# B&R Automation Studio project ProjetoFinalRobotica
Automation Studio 4.1.14.40 SP

## Configuration Config1

CPU 4PP481.1043-B5, AutomationRuntime E3.10, Build 4.1.2, Vc V4.15.9

### Task classes (Cpu.sw)
```
Cyclic#1 (cycle 10000 us, tolerance 10000 us):
  NewProgram <- NewProgram.prg
VcDataObjects: Visu <- Visualisation.Visu.dob
Binaries: arial, Visu02, vccovl, vcdsloc, vcfntttf, vcbclass, vcrt, Visu03, vcfile, vcdsint, vccbtn, vcgclass, vcpdsw, vcshared, vcalarm, arialbd, vcpfpp30, vcmgr, vcpdpp30, Visu01, vctcal, vcpk, vcpfmtcx, vcptelo, ashwd, sysconf, asfw, arconfig, iomap, arialxsr, vcctrend, vccline, vccshape, vccbmp, vcclbox, vccalarm, vccstr, vcchspot, vccgauge, vccurl, vccslider, vccnum, vccdt, vcxml, vccbar, vcchtml, vcctext
Libraries: standard, dataobj, vcresman, fileio, astime, asieccon, AsUDP, Runtime
```

### Hardware
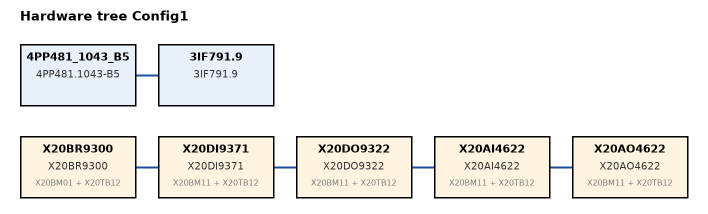
```
3IF791.9 : 3IF791.9 v1.0.0.1  [SS -> 4PP481_1043_B5.SS1]
4PP481_1043_B5 : 4PP481.1043-B5 v1.0.0.0
  Connector IF5:
    ActivateDevice = 1
    Mode = Manual
    InternetAddress = 192.168.0.70
  Cyclic1Duration = 10000
  Cyclic1Tolerance = 10000
  Cyclic2Duration = 20000
  Cyclic2Tolerance = 20000
  Cyclic3Duration = 50000
  Cyclic3Tolerance = 50000
  Cyclic4Duration = 100000
  Cyclic4Tolerance = 100000
  Cyclic5Duration = 200000
  Cyclic5Tolerance = 200000
  Cyclic6Duration = 500000
  Cyclic6Tolerance = 500000
  Cyclic7Duration = 1000000
  Cyclic7Tolerance = 1000000
  Cyclic8Duration = 10000
  Cyclic8Tolerance = 30000000
  VcObjectName = Visu
  KeyMappingFile = VC\4PP481_1043_B5.dis
X20AI4622 : X20AI4622 v1.0.2.0  [SS1 -> X20TB12c.SS; SL -> X20BM11b.SL1]
X20AO4622 : X20AO4622 v1.0.4.0  [SS1 -> X20TB12e.SS; SL -> X20BM11c.SL1]
X20BM01 : X20BM01 v1.0.0.1
X20BM11 : X20BM11 v1.0.0.0  [X2X1 -> X20BM01.X2X2]
X20BM11a : X20BM11 v1.0.0.0  [X2X1 -> X20BM11.X2X2]
X20BM11b : X20BM11 v1.0.0.0  [X2X1 -> X20BM11a.X2X2]
X20BM11c : X20BM11 v1.0.0.0  [X2X1 -> X20BM11b.X2X2]
X20BR9300 : X20BR9300 v1.0.2.4  [SS1 -> X20TB12.SS; SL -> X20BM01.SL1; X2X1 -> 3IF791.9.IF1]
X20DI9371 : X20DI9371 v1.0.1.1  [SS1 -> X20TB12a.SS; SL -> X20BM11.SL1]
X20DO9322 : X20DO9322 v1.0.2.2  [SS1 -> X20TB12b.SS; SL -> X20BM11a.SL1]
X20TB12 : X20TB12 v1.0.0.0
X20TB12a : X20TB12 v1.0.0.0
X20TB12b : X20TB12 v1.0.0.0
X20TB12c : X20TB12 v1.0.0.0
X20TB12e : X20TB12 v1.0.0.0
```

### IoMap.iom - 4PP481_1043_B5/IoMap.iom
```iecst
(********************************************************************
 * COPYRIGHT --
 ********************************************************************
 * File: IoMap.iom
 * Author: supervisorio
 * Created: February 20, 2025
 ********************************************************************
 * IO mapping file
 ********************************************************************)
VAR_CONFIG
	::NewProgram:Jaka_DI3 AT %QX."X20DO9322".DigitalOutput01;
	::NewProgram:Jaka_DI2 AT %QX."X20DO9322".DigitalOutput02;
	::NewProgram:Jaka_DI1 AT %QX."X20DO9322".DigitalOutput03;
	::NewProgram:Staubli_DI12 AT %QX."X20DO9322".DigitalOutput05;
	::NewProgram:Staubli_DI13 AT %QX."X20DO9322".DigitalOutput06;
	::NewProgram:Staubli_DI14 AT %QX."X20DO9322".DigitalOutput07;
	::NewProgram:Staubli_DI15 AT %QX."X20DO9322".DigitalOutput08;
	::NewProgram:Esteira_StaubliJaka AT %QX."X20DO9322".DigitalOutput11;
	::NewProgram:Esteira_JakaStaubli AT %QX."X20DO9322".DigitalOutput12;
	::NewProgram:Jaka_DO7 AT %IX."X20DI9371".DigitalInput01;
	::NewProgram:Jaka_DO6 AT %IX."X20DI9371".DigitalInput02;
	::NewProgram:Jaka_DO5 AT %IX."X20DI9371".DigitalInput03;
	::NewProgram:Staubli_DO4 AT %IX."X20DI9371".DigitalInput05;
	::NewProgram:Staubli_DO5 AT %IX."X20DI9371".DigitalInput06;
	::NewProgram:Staubli_DO6 AT %IX."X20DI9371".DigitalInput07;
	::NewProgram:Staubli_DO7 AT %IX."X20DI9371".DigitalInput08;
	::NewProgram:Sensor_Staubli AT %IX."X20DI9371".DigitalInput09;
	::NewProgram:Sensor_Jaka AT %IX."X20DI9371".DigitalInput10;
	::NewProgram:Emergencia AT %IX."X20DI9371".DigitalInput12;
END_VAR
```

## Logical view

Binary libraries used (declarations not repeated): operator, runtime, astime, AsIecCon, standard, AsUDP

### Global.typ - Global data types
```iecst
(********************************************************************
 * COPYRIGHT --
 ********************************************************************
 * File: Global.typ
 * Author: supervisorio
 * Created: February 20, 2025
 ********************************************************************
 * Global data types of project CLP_ROBO
 ********************************************************************)

TYPE
	feeder_status_typ : 	STRUCT
		power : BOOL;
		home : BOOL;
		axisErrorNumber : UINT;
		axisErrorText : STRING[255];
	END_STRUCT;
	feeder_cmd_typ : 	STRUCT
		requestToPut : BOOL;
	END_STRUCT;
	feeder_typ : 	STRUCT
		cmd : feeder_cmd_typ;
		status : feeder_status_typ;
	END_STRUCT;
	main_status_money_typ : 	STRUCT
		changedMoney : REAL;
		cent1 : USINT;
		cent2 : USINT;
		cent5 : USINT;
		cent10 : USINT;
		cent20 : USINT;
		cent50 : USINT;
		euro1 : UDINT;
		euro2 : UDINT;
	END_STRUCT;
	main_status_progress_typ : 	STRUCT
		total : REAL;
		current : REAL;
	END_STRUCT;
	main_status_typ : 	STRUCT
		money : main_status_money_typ;
		progressStep : USINT;
		curPage : UINT;
		curLanguage : UINT;
		startProgressStep : USINT;
	END_STRUCT;
	main_par_recipe_typ : 	STRUCT
		price : REAL;
		setTemp : REAL;
		milk : REAL;
		sugar : REAL;
		coffee : REAL;
		water : REAL;
	END_STRUCT;
	main_par_typ : 	STRUCT
		coffeeType : SINT;
		givenMoney : REAL;
		recipe : main_par_recipe_typ;
	END_STRUCT;
	main_cmd_typ : 	STRUCT
		switchOnOff : BOOL;
		errorAck : BOOL;
		start : BOOL;
		vis : main_cmd_vis_typ;
	END_STRUCT;
	main_cmd_vis_typ : 	STRUCT
		newPage : UINT;
		startFlag : BOOL;
		startButtonColor : UINT;
		waterTempColor : UINT;
		messageColor : UINT;
		messageIndex : USINT;
		euro2hidden : UINT;
		euro1hidden : UINT;
		cent50hidden : UINT;
		cent20hidden : UINT;
		cent10hidden : UINT;
		cent5hidden : UINT;
		cent2hidden : UINT;
		cent1hidden : UINT;
		newLanguage : UINT;
	END_STRUCT;
	main_typ : 	STRUCT
		cmd : main_cmd_typ;
		par : main_par_typ;
		status : main_status_typ;
	END_STRUCT;
	conveyor_typ : 	STRUCT
		status : conveyor_status_typ;
	END_STRUCT;
	conveyor_status_typ : 	STRUCT
		power : BOOL;
		home : BOOL;
		axisErrorNumber : UINT;
		axisErrorText : STRING[255];
		readyToTake : BOOL;
	END_STRUCT;
	brewing_par_typ : 	STRUCT
		coffeeType : USINT;
	END_STRUCT;
	brewing_cmd_typ : 	STRUCT
		start : BOOL;
	END_STRUCT;
	brewing_status_typ : 	STRUCT
		done : BOOL;
		sBrewingStep : UINT;
		brewingStepText : STRING[64];
	END_STRUCT;
	brewing_typ : 	STRUCT
		cmd : brewing_cmd_typ;
		par : brewing_par_typ;
		status : brewing_status_typ;
	END_STRUCT;
	heating_status_typ : 	STRUCT
		setTempOK : BOOL;
		actTemp : REAL;
	END_STRUCT;
	heating_cmd_typ : 	STRUCT
		start : BOOL;
		updatePIDpar : BOOL;
	END_STRUCT;
	heating_typ : 	STRUCT
		cmd : heating_cmd_typ;
		status : heating_status_typ;
	END_STRUCT;
END_TYPE
```

### Package Logical/Libraries - Global libraries

- Visualisation Logical/Visualisation (not shown)

### Program Logical/NewProgram (IEC) - Program

#### NewProgramCyclic.st - Cyclic code
```iecst
(********************************************************************
 * COPYRIGHT --
 ********************************************************************
 * PROGRAM: NewProgram
 * File: NewProgramCyclic.st
 * Author: supervisorio
 * Created: May 29, 2026
 ********************************************************************
 * Whiteboard application (docs/whiteboard-application.md):
 *   1. Jaka puts the plate (NUM_PECAS parts in its holes) on the conveyor.
 *   2. The conveyor brings the plate TO the Staubli.
 *   3. Staubli puts the plate on its table AND the parts on the board.
 *   4. Staubli picks the marker from its table, draws a square around
 *      each part AND puts the marker back.
 * NUM_PECAS (NewProgram.var) is 1 FOR now: one part, one square.
 * Every robot task uses a four-phase handshake (no timers):
 *   PLC sets CMD -> robot sets DONE -> PLC clears CMD -> robot clears DONE.
 * One run per press OF the start button: Ligar is cleared at the end
 * OF the cycle AND on E-stop.
 ********************************************************************)
PROGRAM _CYCLIC

	TmrPulso(IN := Ligar AND Emergencia, PT := T#1s);
	TmrDI12(IN := Etapa = 2, PT := T#1s);

	IF Ligar AND Emergencia THEN

		Jaka_DI2 := NOT TmrPulso.Q;		//Pulse: ON for the first 1 s of the cycle, then OFF
		Staubli_DI13 := NOT TmrPulso.Q;
		LIGA_JAKA := TRUE;

		CASE Etapa OF

			0: (* Start *)
				PlacaNaEsteira := FALSE;
				PlacaChegou := FALSE;
				PecasNoQuadro := FALSE;
				CicloConcluido := FALSE;
				iPecasNoQuadro := 0;
				iQuadrados := 0;
				iTempoCiclo_s := 0;
				Jaka_DI3 := TRUE;						//CMD Jaka: put the plate on the conveyor
				Etapa := 1;

			1: (* Plate to the Staubli *)
				IF Jaka_DO7 = TRUE THEN
					//Jaka_DI3 := FALSE;					//Jaka done: plate on the conveyor
					PlacaNaEsteira := TRUE;
					Esteira_JakaStaubli := TRUE;
					Jaka_DI2 := FALSE;	//Carry the plate to the Staubli
				END_IF;

				IF Esteira_JakaStaubli AND Sensor_Staubli THEN
					Esteira_JakaStaubli := FALSE;		//Plate arrived
					PlacaChegou := TRUE;
				END_IF;

				//Wait for the Jaka to clear DONE
				IF PlacaChegou AND NOT Jaka_DO7 THEN
					Etapa := 2;
				END_IF;

			2: (* Staubli: plate on the table, parts on the board *)
				Staubli_DI12 := NOT TmrDI12.Q;			//CMD Staubli: plate to the table, parts to the board
				IF Staubli_DO4 THEN
					Staubli_DI12 := FALSE;				//Staubli done: parts on the board
					PecasNoQuadro := TRUE;
					iPecasNoQuadro := NUM_PECAS;
					Etapa := 3;
				END_IF;

			3: (* Wait for the Staubli to clear DONE *)
				IF NOT Staubli_DO4 THEN
					Etapa := 4;
				END_IF;

			4: (* Staubli: pick the marker, draw the squares, put the marker back *)
				Staubli_DI14 := TRUE;					//CMD Staubli: pick the marker and draw
				IF Staubli_DO5 THEN
					Staubli_DI14 := FALSE;				//Staubli done: squares drawn, marker stored
					iQuadrados := NUM_PECAS;
					Etapa := 5;
				END_IF;

			5: (* Finish: wait for the Staubli to clear DONE *)
				IF NOT Staubli_DO5 THEN
					iContador := iContador + 1;			//Completed cycles
					CicloConcluido := TRUE;
					Ligar := FALSE;						//One run per start; press Ligar again for the next
					Etapa := 0;
				END_IF;

		END_CASE;

	ELSE
		//Stop or E-stop: every command and enable goes FALS
		LIGA_JAKA := FALSE;
		Jaka_DI1 := FALSE;
		Jaka_DI2 := FALSE;
		Jaka_DI3 := FALSE;
		Staubli_DI12 := FALSE;
		Staubli_DI13 := FALSE;
		Staubli_DI14 := FALSE;
		Staubli_DI15 := FALSE;
		Esteira_JakaStaubli := FALSE;
		Esteira_StaubliJaka := FALSE;
		IF NOT Emergencia THEN
			Ligar := FALSE;							//Releasing the E-stop must not restart the cell
		END_IF;
		Etapa := 0;

		//Reset the process state too, so the HMI colors, counters and progress go back to "waiting".
		//Skipped right after a finished cycle: CicloConcluido stays TRUE until the next start,
		//so the "done" state and the cycle time stay on screen.
		IF NOT CicloConcluido THEN
			PlacaNaEsteira := FALSE;
			PlacaChegou := FALSE;
			PecasNoQuadro := FALSE;
			iPecasNoQuadro := 0;
			iQuadrados := 0;
			iTempoCiclo_s := 0;
		END_IF;
	END_IF;

	//Progress counters from the robots' optional pulses (Staubli DO6 = part placed, DO7 = square drawn)
	PulsoPeca(CLK := Staubli_DO6);
	IF PulsoPeca.Q AND Etapa = 2 AND iPecasNoQuadro < NUM_PECAS THEN
		iPecasNoQuadro := iPecasNoQuadro + 1;
	END_IF;
	PulsoQuadrado(CLK := Staubli_DO7);
	IF PulsoQuadrado.Q AND Etapa = 4 AND iQuadrados < NUM_PECAS THEN
		iQuadrados := iQuadrados + 1;
	END_IF;

	//Cycle time (kept on screen after the cycle ends)
	TempoCiclo(IN := Etapa > 0, PT := T#30m);
	IF Etapa > 0 THEN
		iTempoCiclo_s := DINT_TO_INT(TIME_TO_DINT(TempoCiclo.ET) / 1000);
	END_IF;

	//Where the plate is: 0 = Jaka, 1 = conveyor, 2 = Staubli
	IF PlacaChegou THEN
		iPlaca := 2;
	ELSIF PlacaNaEsteira THEN
		iPlaca := 1;
	ELSE
		iPlaca := 0;
	END_IF;

	//HMI colors (palette index): COR_ESPERA = waiting, COR_ANDAMENTO = running, COR_FEITO = done
	IF PlacaNaEsteira THEN iCorJaka := COR_FEITO; ELSIF Jaka_DI3 THEN iCorJaka := COR_ANDAMENTO; ELSE iCorJaka := COR_ESPERA; END_IF;
	IF PlacaChegou THEN iCorEsteira := COR_FEITO; ELSIF Esteira_JakaStaubli THEN iCorEsteira := COR_ANDAMENTO; ELSE iCorEsteira := COR_ESPERA; END_IF;
	IF PecasNoQuadro THEN iCorPecas := COR_FEITO; ELSIF Staubli_DI12 THEN iCorPecas := COR_ANDAMENTO; ELSE iCorPecas := COR_ESPERA; END_IF;
	IF CicloConcluido OR Etapa = 5 THEN iCorDesenho := COR_FEITO; ELSIF Etapa = 4 THEN iCorDesenho := COR_ANDAMENTO; ELSE iCorDesenho := COR_ESPERA; END_IF;
	IF CicloConcluido THEN iCorConcluido := COR_FEITO; ELSIF Etapa = 5 THEN iCorConcluido := COR_ANDAMENTO; ELSE iCorConcluido := COR_ESPERA; END_IF;

	//Whiteboard (one part and its square on the HMI)
	IF iPecasNoQuadro >= 1 THEN iCorPeca := COR_PECA; ELSE iCorPeca := COR_VAZIO; END_IF;
	IF iQuadrados >= 1 THEN iCorQuadrado := COR_TINTA; ELSE iCorQuadrado := COR_QUADRO; END_IF;

	IF iPlaca = 0 THEN iCorPlacaJaka := COR_FEITO; ELSE iCorPlacaJaka := COR_ESPERA; END_IF;
	IF iPlaca = 1 THEN iCorPlacaEsteira := COR_FEITO; ELSE iCorPlacaEsteira := COR_ESPERA; END_IF;
	IF iPlaca = 2 THEN iCorPlacaStaubli := COR_FEITO; ELSE iCorPlacaStaubli := COR_ESPERA; END_IF;

	iProgresso := iPecasNoQuadro + iQuadrados;	//0..2*NUM_PECAS on the progress bar

	//Digital twin: send the I/O state to the bridge PC (TwinSender.st)
	TwinSender;

END_PROGRAM
```

#### TwinSender.st - Digital twin UDP sender (action)
```iecst
(********************************************************************
 * COPYRIGHT --
 ********************************************************************
 * Program: NewProgram
 * File: TwinSender.st
 ********************************************************************
 * Digital twin: sends the I/O state to the bridge PC over UDP.
 * Called once per scan at the end of _CYCLIC.
 * Packet layout: docs/publishing-plan/02-plc-udp-sender.md
 * Needs the AsUDP library (Logical View > Libraries > Add Object).
 * Send errors are only counted: the cell must never depend on the
 * bridge PC being present.
 ********************************************************************)
ACTION TwinSender:

	(* Bytes 0..11: X20DI9371 channels 1..12 *)
	TwinPacket[0]  := BOOL_TO_USINT(Jaka_DO7);
	TwinPacket[1]  := BOOL_TO_USINT(Jaka_DO6);
	TwinPacket[2]  := BOOL_TO_USINT(Jaka_DO5);
	TwinPacket[4]  := BOOL_TO_USINT(Staubli_DO4);
	TwinPacket[5]  := BOOL_TO_USINT(Staubli_DO5);
	TwinPacket[6]  := BOOL_TO_USINT(Staubli_DO6);
	TwinPacket[7]  := BOOL_TO_USINT(Staubli_DO7);
	TwinPacket[8]  := BOOL_TO_USINT(Sensor_Staubli);
	TwinPacket[9]  := BOOL_TO_USINT(Sensor_Jaka);
	TwinPacket[11] := BOOL_TO_USINT(Emergencia);

	(* Bytes 12..23: X20DO9322 channels 1..12 *)
	TwinPacket[12] := BOOL_TO_USINT(Jaka_DI3);
	TwinPacket[13] := BOOL_TO_USINT(LIGA_JAKA);
	TwinPacket[14] := BOOL_TO_USINT(Jaka_DI1);
	TwinPacket[16] := BOOL_TO_USINT(Staubli_DI12);
	TwinPacket[17] := BOOL_TO_USINT(Staubli_DI13);
	TwinPacket[18] := BOOL_TO_USINT(Staubli_DI14);
	TwinPacket[19] := BOOL_TO_USINT(Staubli_DI15);
	TwinPacket[22] := BOOL_TO_USINT(Esteira_StaubliJaka);
	TwinPacket[23] := BOOL_TO_USINT(Esteira_JakaStaubli);

	(* Bytes 24..26: sequence state. Byte 27 (counter) is set when sending. *)
	TwinPacket[24] := INT_TO_USINT(Etapa);
	TwinPacket[25] := INT_TO_USINT(iContador);
	TwinPacket[26] := BOOL_TO_USINT(Ligar);

	CASE TwinState OF

		0: (* open the UDP socket *)
			TwinOpen(enable := TRUE, pIfAddr := 0, port := TwinLocalPort, options := 0);
			IF TwinOpen.status = ERR_OK THEN
				TwinState := 1;
			ELSIF TwinOpen.status <> ERR_FUB_BUSY THEN
				TwinOpenErr := TwinOpen.status;     // erro real, antes de desligar o bloco
				TwinOpen(enable := FALSE);
				TwinState := 3;
			END_IF;

		1: (* wait for the next period *)
			TwinTimer(IN := TRUE, PT := T#200ms);
			IF TwinTimer.Q THEN
				TwinTimer(IN := FALSE);
				TwinSeq := TwinSeq + 1;
				TwinPacket[27] := TwinSeq;
				TwinState := 2;
			END_IF;

		2: (* send; keep calling while busy *)
			TwinSend(enable := TRUE, ident := TwinOpen.ident, pHost := ADR(TwinHost), port := TwinPort,
				pData := ADR(TwinPacket), datalen := SIZEOF(TwinPacket), flags := 0);
			IF TwinSend.status <> ERR_FUB_BUSY THEN
				IF TwinSend.status <> ERR_OK THEN
					TwinSendErrors := TwinSendErrors + 1;
				END_IF;
				TwinSend(enable := FALSE);
				TwinState := 1;
			END_IF;

		3: (* opening failed: try again in 5 s *)
			TwinTimer(IN := TRUE, PT := T#5s);
			IF TwinTimer.Q THEN
				TwinTimer(IN := FALSE);
				TwinState := 0;
			END_IF;

	END_CASE;

END_ACTION
```

#### NewProgram.var - Local variables
```iecst
(********************************************************************
 * COPYRIGHT --
 ********************************************************************
 * Program: NewProgram
 * File: NewProgram.var
 * Author: supervisorio
 * Created: May 29, 2026
 ********************************************************************
 * Local variables of program NewProgram
 ********************************************************************)
(* I/O, mapped in IoMap.iom (Table I of the cell handout) *)
VAR
	Emergencia : BOOL;
	Jaka_DO7 : BOOL; (*DONE: plate on the conveyor*)
	Jaka_DO6 : BOOL; (*spare*)
	Jaka_DO5 : BOOL; (*pulse: plate gripped (twin only)*)
	Jaka_DI3 : BOOL; (*CMD: put the plate on the conveyor*)
	Jaka_DI2 : BOOL; (*enable*)
	Jaka_DI1 : BOOL; (*spare*)
	Staubli_DO4 : BOOL; (*DONE: plate on the table, part on the board*)
	Staubli_DO5 : BOOL; (*DONE: square drawn, marker stored*)
	Staubli_DO6 : BOOL; (*pulse: one part placed*)
	Staubli_DO7 : BOOL; (*pulse: one square drawn*)
	Staubli_DI12 : BOOL; (*CMD: plate to the table, part to the board*)
	Staubli_DI13 : BOOL; (*enable*)
	Staubli_DI14 : BOOL; (*CMD: pick the marker and draw*)
	Staubli_DI15 : BOOL; (*spare*)
	Esteira_StaubliJaka : BOOL; (*spare*)
	Esteira_JakaStaubli : BOOL; (*carries the plate to the Staubli*)
	Sensor_Jaka : BOOL;
	Sensor_Staubli : BOOL;
END_VAR
(* Sequence *)
VAR CONSTANT
	NUM_PECAS : INT := 1; (*parts on the plate per run; one square is drawn around each*)
END_VAR
VAR
	Ligar : BOOL; (*start request from the HMI, cleared at the end of the cycle*)
	Etapa : INT; (*0 idle, 1 plate to Staubli, 2 parts to board, 3 wait, 4 drawing, 5 finishing*)
	PlacaNaEsteira : BOOL;
	PlacaChegou : BOOL;
	PecasNoQuadro : BOOL;
	CicloConcluido : BOOL;
	iContador : INT; (*completed cycles*)
	PulsoPeca : R_TRIG;
	PulsoQuadrado : R_TRIG;
	TempoCiclo : TON;
END_VAR
(* HMI (Init_Page) *)
VAR
	iPecasNoQuadro : INT; (*0..NUM_PECAS*)
	iQuadrados : INT; (*0..NUM_PECAS*)
	iTempoCiclo_s : INT; (*seconds*)
	iPlaca : INT; (*plate: 0 Jaka, 1 conveyor, 2 Staubli*)
	iProgresso : INT; (*0..2*NUM_PECAS*)
	iCorJaka : INT;
	iCorEsteira : INT;
	iCorPecas : INT;
	iCorDesenho : INT;
	iCorConcluido : INT;
	iCorPeca : INT;
	iCorQuadrado : INT;
	iCorPlacaJaka : INT;
	iCorPlacaEsteira : INT;
	iCorPlacaStaubli : INT;
END_VAR
(* HMI palette indexes (Palette.vcr) *)
VAR CONSTANT
	COR_ESPERA : INT := 250; (*light grey: waiting*)
	COR_ANDAMENTO : INT := 46; (*yellow: running*)
	COR_FEITO : INT := 155; (*green: done*)
	COR_ALARME : INT := 51; (*red*)
	COR_PECA : INT := 204; (*blue: part on the board*)
	COR_VAZIO : INT := 252; (*very light grey: empty slot*)
	COR_TINTA : INT := 0; (*black: square drawn*)
	COR_QUADRO : INT := 15; (*white: whiteboard*)
END_VAR
(* Digital twin UDP sender (TwinSender.st). Set TwinHost to the IP of the bridge PC. *)
VAR
	TwinHost : STRING[15] := '192.168.0.100'; (*IP of the bridge PC on the cell network*)
	TwinPort : UINT := 5005; (*UDP port the bridge listens on*)
	TwinLocalPort : UINT := 5006; (*local UDP port on the PLC*)
	TwinOpen : UdpOpen;
	TwinSend : UdpSend;
	TwinTimer : TON;
	TwinPacket : ARRAY[0..27] OF USINT;
	TwinSeq : USINT;
	TwinState : USINT;
	TwinSendErrors : UDINT; (*failed sends, for diagnosis only*)
	TwinOpenErr : UDINT;
	TmrPulso : TON;
	TmrDI12 : TON;
	LIGA_JAKA : BOOL;
END_VAR
```
